KUKA KRL program: MAIN_1.src

&ACCESS RVP
&REL 1
&PARAM TEMPLATE = C:\KRC\Roboter\Template\vorgabe
&PARAM EDITMASK = *
DEF MAIN_1 ( )

; External program calls:
EXT REMOTE_PROG_CALL_171()
EXT PICK_PART_111()
EXT PLACE_PART_112()
EXT EVENT_PROG_START_101()
EXT EVENT_PATH_APPROACH_102()
EXT EVENT_PATH_START_103()
EXT EVENT_PATH_FINISH_105()
EXT EVENT_PATH_RETRACT_106()
EXT EVENT_PROG_FINISH_107()
EXT PROG_1___with_a_very_long_name_and_special_characters()


EXT CLEENING ()
;FOLD INI

;FOLD BASISTECH INI
GLOBAL INTERRUPT DECL 3 WHEN $STOPMESS==TRUE DO IR_STOPM ( )
INTERRUPT ON 3
BAS (#INITMOV,0)
BAS (#VEL_PTP,20)
BAS (#ACC_PTP,20)
;ENDFOLD (BASISTECH INI)

;FOLD SPOTTECH INI
;USERSPOT(#INIT)
;ENDFOLD (SPOTTECH INI)

;FOLD GRIPPERTECH INI
;USER_GRP(0,DUMMY,DUMMY,GDEFAULT)
;ENDFOLD (GRIPPERTECH INI)

;FOLD ARCTECHDIGITAL INI
IF ARC20==TRUE THEN
  A20 (ARC_INI)
  INTERRUPT DECL 6 WHEN $CYCFLAG[3]==FALSE DO A20(TECH_STOP2)
ENDIF
;ENDFOLD (ARCTECHDIGITAL INI)

;FOLD USER INI
;---- Make your modifications here ----

;ENDFOLD (USER INI)

;ENDFOLD (INI)


;FOLD PTP HOME Vel=20 % DEFAULT;%{PE}%R 5.6.13,%MKUKATPBASIS,%CMOVE,%VPTP,%P 1:PTP, 2:HOME, 3:, 5:20, 7:DEFAULT
$BWDSTART=FALSE
PDAT_ACT=PDEFAULT
FDAT_ACT=FHOME
BAS(#PTP_PARAMS,20)
$H_POS=XHOME
PTP XHOME
;ENDFOLD


; Program generated by RoboDK v5.6.9 for RoboDK Industrial on 26/02/2024 09:58:20
; Using nominal kinematics.
;FOLD PTP P1 Vel=100.000 % PDAT1 Tool[1] Base[1];%{PE}%R 5.5.31,%MKUKATPBASIS,%CMOVE,%VPTP,%P 1:PTP, 2:P1, 3:, 5:100.000, 7:PDAT1
$BWDSTART=FALSE
PDAT_ACT=PPDAT1
FDAT_ACT=FP1
BAS(#PTP_PARAMS,100)
PTP XP1 C_PTP
;ENDFOLD

;FOLD PTP P2 Vel=100.000 % PDAT2 Tool[1] Base[1];%{PE}%R 5.5.31,%MKUKATPBASIS,%CMOVE,%VPTP,%P 1:PTP, 2:P2, 3:, 5:100.000, 7:PDAT2
$BWDSTART=FALSE
PDAT_ACT=PPDAT2
FDAT_ACT=FP2
BAS(#PTP_PARAMS,100)
PTP XP2 C_PTP
;ENDFOLD

;FOLD LIN P3 Vel=1.000 m/s CPDAT3 Tool[1] Base[1];%{PE}%R 5.5.0,%MKUKATPA20,%CARC_SWI,%VLIN,%P 1:LIN, 2:P3, 3:, 5:1.000, 7:CPDAT3
$BWDSTART=FALSE
LDAT_ACT=LCPDAT3
FDAT_ACT=FP3
LIN XP3
;ENDFOLD

$OUT[5]=TRUE
$OUT[5]=TRUE
$OUT[5]=0.5
$OUT[5]=true
$ANOUT[5]=TRUE
$ANOUT[5]=TRUE
$ANOUT[5]=0.5
$ANOUT[5]=true
var=val
var=val
WAIT FOR ($IN[5]==TRUE)
WAIT FOR ($IN[5]==TRUE)
WAIT FOR ($IN[5]==0.5)
WAIT FOR ($IN[5]==true)
START_TIMER:
$TIMER_STOP[1]=TRUE
$TIMER_FLAG[1]=FALSE
$TIMER[1]=0.100
$TIMER_STOP[1]=FALSE
WAIT FOR ($IN[5]==TRUE OR $TIMER_FLAG[1])
$TIMER_STOP[1]=TRUE
IF $TIMER_FLAG[1]== TRUE THEN
    HALT ; Timed out!
    GOTO START_TIMER
ENDIF
WAIT FOR (var==val)
START_TIMER:
$TIMER_STOP[1]=TRUE
$TIMER_FLAG[1]=FALSE
$TIMER[1]=0.100
$TIMER_STOP[1]=FALSE
WAIT FOR (var==val OR $TIMER_FLAG[1])
$TIMER_STOP[1]=TRUE
IF $TIMER_FLAG[1]== TRUE THEN
    HALT ; Timed out!
    GOTO START_TIMER
ENDIF
Wait for StrClear($LOOP_MSG[])
$LOOP_CONT = TRUE
$LOOP_MSG[] = "Message"
REMOTE_PROG_CALL_171()
CODE_INSERT_172
; Insert Comment
BASE_DATA[1] = {FRAME: X 719.013,Y -664.003,Z 0.000,A 0.000,B 0.000,C 0.000}
TOOL_DATA[1] = {FRAME: X 129.073,Y 0.000,Z 85.477,A 0.000,B 22.849,C 0.000}
$ACC.ORI1 = 800.00000
$ACC.ORI2 = 800.00000
$VEL.ORI1 = 500.00000
$VEL.ORI2 = 500.00000
$APO.CPTP = 10
$APO.CDIS = 10.000
;FOLD PTP P4 CONT Vel=100.000 % PDAT4 Tool[1] Base[1];%{PE}%R 5.5.31,%MKUKATPBASIS,%CMOVE,%VPTP,%P 1:PTP, 2:P4, 3:C_PTP, 5:100.000, 7:PDAT4
$BWDSTART=FALSE
PDAT_ACT=PPDAT4
FDAT_ACT=FP4
BAS(#PTP_PARAMS,100)
PTP XP4 C_PTP
;ENDFOLD

$ACC.CP = 0.20000
;FOLD LIN P5 Vel=0.100 m/s CPDAT5 Tool[1] Base[1];%{PE}%R 5.5.0,%MKUKATPA20,%CARC_SWI,%VLIN,%P 1:LIN, 2:P5, 3:, 5:0.100, 7:CPDAT5
$BWDSTART=FALSE
LDAT_ACT=LCPDAT5
FDAT_ACT=FP5
LIN XP5
;ENDFOLD

$OUT[5]=TRUE
PICK_PART_111()
$APO.CPTP = 10
$APO.CDIS = 10.000
$ACC.CP = 0.60000
; Linear movement using joint targets is not supported. Change the target type to cartesian or use a joint movement.
;FOLD LIN P6 CONT Vel=0.300 m/s CPDAT6 Tool[1] Base[1];%{PE}%R 5.5.0,%MKUKATPA20,%CARC_SWI,%VLIN,%P 1:LIN, 2:P6, 3:C_DIS, 5:0.300, 7:CPDAT6
$BWDSTART=FALSE
LDAT_ACT=LCPDAT6
FDAT_ACT=FP6
LIN XP6 C_DIS
;ENDFOLD

$ACC.CP = 0.20000
; MoveSearch command not implemented
;FOLD LIN P7 Vel=0.100 m/s CPDAT7 Tool[1] Base[1];%{PE}%R 5.5.0,%MKUKATPA20,%CARC_SWI,%VLIN,%P 1:LIN, 2:P7, 3:, 5:0.100, 7:CPDAT7
$BWDSTART=FALSE
LDAT_ACT=LCPDAT7
FDAT_ACT=FP7
LIN XP7
;ENDFOLD

$OUT[5]=FALSE
PLACE_PART_112()
$APO.CPTP = 10
$APO.CDIS = 10.000
;FOLD LIN P8 CONT Vel=0.100 m/s CPDAT8 Tool[1] Base[1];%{PE}%R 5.5.0,%MKUKATPA20,%CARC_SWI,%VLIN,%P 1:LIN, 2:P8, 3:C_DIS, 5:0.100, 7:CPDAT8
$BWDSTART=FALSE
LDAT_ACT=LCPDAT8
FDAT_ACT=FP8
LIN XP8 C_DIS
;ENDFOLD

BASE_DATA[1] = {FRAME: X 577.670,Y 392.250,Z 0.000,A 38.960,B 0.000,C 0.000}
$APO.CPTP = 25
$APO.CDIS = 25.000
$ACC.ORI1 = 800.00000
$ACC.ORI2 = 800.00000
$VEL.ORI1 = 500.00000
$VEL.ORI2 = 500.00000
$ACC.CP = 0.20000
;FOLD PTP P9 CONT Vel=100.000 % PDAT9 Tool[1] Base[1];%{PE}%R 5.5.31,%MKUKATPBASIS,%CMOVE,%VPTP,%P 1:PTP, 2:P9, 3:C_PTP, 5:100.000, 7:PDAT9
$BWDSTART=FALSE
PDAT_ACT=PPDAT9
FDAT_ACT=FP9
BAS(#PTP_PARAMS,100)
PTP XP9 C_PTP
;ENDFOLD

CIRC {X 430.047,Y 43.774,Z 231.503,A -134.549,B 11.181,C 178.913},{X 109.688,Y -153.222,Z 161.073,A -134.549,B 11.181,C 178.913} C_DIS
; Circular movement using joint targets is not supported. Change the target type to cartesian or use a joint movement.
$ACC.CP = 0.20000
;FOLD LIN P10 Vel=0.100 m/s CPDAT10 Tool[1] Base[1];%{PE}%R 5.5.0,%MKUKATPA20,%CARC_SWI,%VLIN,%P 1:LIN, 2:P10, 3:, 5:0.100, 7:CPDAT10
$BWDSTART=FALSE
LDAT_ACT=LCPDAT10
FDAT_ACT=FP10
LIN XP10
;ENDFOLD

;FOLD PTP P11 Vel=100.000 % PDAT11 Tool[1] Base[1];%{PE}%R 5.5.31,%MKUKATPBASIS,%CMOVE,%VPTP,%P 1:PTP, 2:P11, 3:, 5:100.000, 7:PDAT11
$BWDSTART=FALSE
PDAT_ACT=PPDAT11
FDAT_ACT=FP11
BAS(#PTP_PARAMS,100)
PTP XP11 C_PTP
;ENDFOLD

BASE_DATA[1] = {FRAME: X 0.000,Y 782.714,Z 377.610,A 0.000,B 0.000,C 0.000}
;FOLD PTP P12 Vel=100.000 % PDAT12 Tool[1] Base[1];%{PE}%R 5.5.31,%MKUKATPBASIS,%CMOVE,%VPTP,%P 1:PTP, 2:P12, 3:, 5:100.000, 7:PDAT12
$BWDSTART=FALSE
PDAT_ACT=PPDAT12
FDAT_ACT=FP12
BAS(#PTP_PARAMS,100)
PTP XP12 C_PTP
;ENDFOLD

;FOLD LIN P13 Vel=0.100 m/s CPDAT13 Tool[1] Base[1];%{PE}%R 5.5.0,%MKUKATPA20,%CARC_SWI,%VLIN,%P 1:LIN, 2:P13, 3:, 5:0.100, 7:CPDAT13
$BWDSTART=FALSE
LDAT_ACT=LCPDAT13
FDAT_ACT=FP13
LIN XP13
;ENDFOLD

;FOLD LIN P14 Vel=0.100 m/s CPDAT14 Tool[1] Base[1];%{PE}%R 5.5.0,%MKUKATPA20,%CARC_SWI,%VLIN,%P 1:LIN, 2:P14, 3:, 5:0.100, 7:CPDAT14
$BWDSTART=FALSE
LDAT_ACT=LCPDAT14
FDAT_ACT=FP14
LIN XP14
;ENDFOLD

;FOLD LIN P15 Vel=0.100 m/s CPDAT15 Tool[1] Base[1];%{PE}%R 5.5.0,%MKUKATPA20,%CARC_SWI,%VLIN,%P 1:LIN, 2:P15, 3:, 5:0.100, 7:CPDAT15
$BWDSTART=FALSE
LDAT_ACT=LCPDAT15
FDAT_ACT=FP15
LIN XP15
;ENDFOLD

;FOLD LIN P16 Vel=0.100 m/s CPDAT16 Tool[1] Base[1];%{PE}%R 5.5.0,%MKUKATPA20,%CARC_SWI,%VLIN,%P 1:LIN, 2:P16, 3:, 5:0.100, 7:CPDAT16
$BWDSTART=FALSE
LDAT_ACT=LCPDAT16
FDAT_ACT=FP16
LIN XP16
;ENDFOLD

;FOLD LIN P17 Vel=0.100 m/s CPDAT17 Tool[1] Base[1];%{PE}%R 5.5.0,%MKUKATPA20,%CARC_SWI,%VLIN,%P 1:LIN, 2:P17, 3:, 5:0.100, 7:CPDAT17
$BWDSTART=FALSE
LDAT_ACT=LCPDAT17
FDAT_ACT=FP17
LIN XP17
;ENDFOLD

;FOLD LIN P18 Vel=0.100 m/s CPDAT18 Tool[1] Base[1];%{PE}%R 5.5.0,%MKUKATPA20,%CARC_SWI,%VLIN,%P 1:LIN, 2:P18, 3:, 5:0.100, 7:CPDAT18
$BWDSTART=FALSE
LDAT_ACT=LCPDAT18
FDAT_ACT=FP18
LIN XP18
;ENDFOLD

;FOLD LIN P19 Vel=0.100 m/s CPDAT19 Tool[1] Base[1];%{PE}%R 5.5.0,%MKUKATPA20,%CARC_SWI,%VLIN,%P 1:LIN, 2:P19, 3:, 5:0.100, 7:CPDAT19
$BWDSTART=FALSE
LDAT_ACT=LCPDAT19
FDAT_ACT=FP19
LIN XP19
;ENDFOLD

;FOLD PTP P20 Vel=100.000 % PDAT20 Tool[1] Base[1];%{PE}%R 5.5.31,%MKUKATPBASIS,%CMOVE,%VPTP,%P 1:PTP, 2:P20, 3:, 5:100.000, 7:PDAT20
$BWDSTART=FALSE
PDAT_ACT=PPDAT20
FDAT_ACT=FP20
BAS(#PTP_PARAMS,100)
PTP XP20 C_PTP
;ENDFOLD

EVENT_PROG_START_101()
$APO.CPTP = 1
$APO.CDIS = 1.000
BASE_DATA[1] = {FRAME: X 13.637,Y -840.080,Z 0.000,A -90.000,B 0.000,C 0.000}
; Show Tool 1
;FOLD PTP P21 CONT Vel=100.000 % PDAT21 Tool[1] Base[1];%{PE}%R 5.5.31,%MKUKATPBASIS,%CMOVE,%VPTP,%P 1:PTP, 2:P21, 3:C_PTP, 5:100.000, 7:PDAT21
$BWDSTART=FALSE
PDAT_ACT=PPDAT21
FDAT_ACT=FP21
BAS(#PTP_PARAMS,100)
PTP XP21 C_PTP
;ENDFOLD

EVENT_PATH_APPROACH_102()
;FOLD LIN P22 CONT Vel=1.000 m/s CPDAT22 Tool[1] Base[1];%{PE}%R 5.5.0,%MKUKATPA20,%CARC_SWI,%VLIN,%P 1:LIN, 2:P22, 3:C_DIS, 5:1.000, 7:CPDAT22
$BWDSTART=FALSE
LDAT_ACT=LCPDAT22
FDAT_ACT=FP22
LIN XP22 C_DIS
;ENDFOLD

;FOLD LIN P23 CONT Vel=1.000 m/s CPDAT23 Tool[1] Base[1];%{PE}%R 5.5.0,%MKUKATPA20,%CARC_SWI,%VLIN,%P 1:LIN, 2:P23, 3:C_DIS, 5:1.000, 7:CPDAT23
$BWDSTART=FALSE
LDAT_ACT=LCPDAT23
FDAT_ACT=FP23
LIN XP23 C_DIS
;ENDFOLD

EVENT_PATH_START_103()
;FOLD LIN P24 CONT Vel=0.050 m/s CPDAT24 Tool[1] Base[1];%{PE}%R 5.5.0,%MKUKATPA20,%CARC_SWI,%VLIN,%P 1:LIN, 2:P24, 3:C_DIS, 5:0.050, 7:CPDAT24
$BWDSTART=FALSE
LDAT_ACT=LCPDAT24
FDAT_ACT=FP24
LIN XP24 C_DIS
;ENDFOLD

;FOLD LIN P25 CONT Vel=0.050 m/s CPDAT25 Tool[1] Base[1];%{PE}%R 5.5.0,%MKUKATPA20,%CARC_SWI,%VLIN,%P 1:LIN, 2:P25, 3:C_DIS, 5:0.050, 7:CPDAT25
$BWDSTART=FALSE
LDAT_ACT=LCPDAT25
FDAT_ACT=FP25
LIN XP25 C_DIS
;ENDFOLD

;FOLD LIN P26 CONT Vel=0.050 m/s CPDAT26 Tool[1] Base[1];%{PE}%R 5.5.0,%MKUKATPA20,%CARC_SWI,%VLIN,%P 1:LIN, 2:P26, 3:C_DIS, 5:0.050, 7:CPDAT26
$BWDSTART=FALSE
LDAT_ACT=LCPDAT26
FDAT_ACT=FP26
LIN XP26 C_DIS
;ENDFOLD

;FOLD LIN P27 CONT Vel=0.050 m/s CPDAT27 Tool[1] Base[1];%{PE}%R 5.5.0,%MKUKATPA20,%CARC_SWI,%VLIN,%P 1:LIN, 2:P27, 3:C_DIS, 5:0.050, 7:CPDAT27
$BWDSTART=FALSE
LDAT_ACT=LCPDAT27
FDAT_ACT=FP27
LIN XP27 C_DIS
;ENDFOLD

;FOLD LIN P28 CONT Vel=0.050 m/s CPDAT28 Tool[1] Base[1];%{PE}%R 5.5.0,%MKUKATPA20,%CARC_SWI,%VLIN,%P 1:LIN, 2:P28, 3:C_DIS, 5:0.050, 7:CPDAT28
$BWDSTART=FALSE
LDAT_ACT=LCPDAT28
FDAT_ACT=FP28
LIN XP28 C_DIS
;ENDFOLD

;FOLD LIN P29 CONT Vel=0.050 m/s CPDAT29 Tool[1] Base[1];%{PE}%R 5.5.0,%MKUKATPA20,%CARC_SWI,%VLIN,%P 1:LIN, 2:P29, 3:C_DIS, 5:0.050, 7:CPDAT29
$BWDSTART=FALSE
LDAT_ACT=LCPDAT29
FDAT_ACT=FP29
LIN XP29 C_DIS
;ENDFOLD

;FOLD LIN P30 CONT Vel=0.050 m/s CPDAT30 Tool[1] Base[1];%{PE}%R 5.5.0,%MKUKATPA20,%CARC_SWI,%VLIN,%P 1:LIN, 2:P30, 3:C_DIS, 5:0.050, 7:CPDAT30
$BWDSTART=FALSE
LDAT_ACT=LCPDAT30
FDAT_ACT=FP30
LIN XP30 C_DIS
;ENDFOLD

;FOLD LIN P31 CONT Vel=0.050 m/s CPDAT31 Tool[1] Base[1];%{PE}%R 5.5.0,%MKUKATPA20,%CARC_SWI,%VLIN,%P 1:LIN, 2:P31, 3:C_DIS, 5:0.050, 7:CPDAT31
$BWDSTART=FALSE
LDAT_ACT=LCPDAT31
FDAT_ACT=FP31
LIN XP31 C_DIS
;ENDFOLD

;FOLD LIN P32 CONT Vel=0.050 m/s CPDAT32 Tool[1] Base[1];%{PE}%R 5.5.0,%MKUKATPA20,%CARC_SWI,%VLIN,%P 1:LIN, 2:P32, 3:C_DIS, 5:0.050, 7:CPDAT32
$BWDSTART=FALSE
LDAT_ACT=LCPDAT32
FDAT_ACT=FP32
LIN XP32 C_DIS
;ENDFOLD

;FOLD LIN P33 CONT Vel=0.050 m/s CPDAT33 Tool[1] Base[1];%{PE}%R 5.5.0,%MKUKATPA20,%CARC_SWI,%VLIN,%P 1:LIN, 2:P33, 3:C_DIS, 5:0.050, 7:CPDAT33
$BWDSTART=FALSE
LDAT_ACT=LCPDAT33
FDAT_ACT=FP33
LIN XP33 C_DIS
;ENDFOLD

;FOLD LIN P34 CONT Vel=0.050 m/s CPDAT34 Tool[1] Base[1];%{PE}%R 5.5.0,%MKUKATPA20,%CARC_SWI,%VLIN,%P 1:LIN, 2:P34, 3:C_DIS, 5:0.050, 7:CPDAT34
$BWDSTART=FALSE
LDAT_ACT=LCPDAT34
FDAT_ACT=FP34
LIN XP34 C_DIS
;ENDFOLD

;FOLD LIN P35 CONT Vel=0.050 m/s CPDAT35 Tool[1] Base[1];%{PE}%R 5.5.0,%MKUKATPA20,%CARC_SWI,%VLIN,%P 1:LIN, 2:P35, 3:C_DIS, 5:0.050, 7:CPDAT35
$BWDSTART=FALSE
LDAT_ACT=LCPDAT35
FDAT_ACT=FP35
LIN XP35 C_DIS
;ENDFOLD

;FOLD LIN P36 CONT Vel=0.050 m/s CPDAT36 Tool[1] Base[1];%{PE}%R 5.5.0,%MKUKATPA20,%CARC_SWI,%VLIN,%P 1:LIN, 2:P36, 3:C_DIS, 5:0.050, 7:CPDAT36
$BWDSTART=FALSE
LDAT_ACT=LCPDAT36
FDAT_ACT=FP36
LIN XP36 C_DIS
;ENDFOLD

;FOLD LIN P37 CONT Vel=0.050 m/s CPDAT37 Tool[1] Base[1];%{PE}%R 5.5.0,%MKUKATPA20,%CARC_SWI,%VLIN,%P 1:LIN, 2:P37, 3:C_DIS, 5:0.050, 7:CPDAT37
$BWDSTART=FALSE
LDAT_ACT=LCPDAT37
FDAT_ACT=FP37
LIN XP37 C_DIS
;ENDFOLD

;FOLD LIN P38 CONT Vel=0.050 m/s CPDAT38 Tool[1] Base[1];%{PE}%R 5.5.0,%MKUKATPA20,%CARC_SWI,%VLIN,%P 1:LIN, 2:P38, 3:C_DIS, 5:0.050, 7:CPDAT38
$BWDSTART=FALSE
LDAT_ACT=LCPDAT38
FDAT_ACT=FP38
LIN XP38 C_DIS
;ENDFOLD

;FOLD LIN P39 CONT Vel=0.050 m/s CPDAT39 Tool[1] Base[1];%{PE}%R 5.5.0,%MKUKATPA20,%CARC_SWI,%VLIN,%P 1:LIN, 2:P39, 3:C_DIS, 5:0.050, 7:CPDAT39
$BWDSTART=FALSE
LDAT_ACT=LCPDAT39
FDAT_ACT=FP39
LIN XP39 C_DIS
;ENDFOLD

;FOLD LIN P40 CONT Vel=0.050 m/s CPDAT40 Tool[1] Base[1];%{PE}%R 5.5.0,%MKUKATPA20,%CARC_SWI,%VLIN,%P 1:LIN, 2:P40, 3:C_DIS, 5:0.050, 7:CPDAT40
$BWDSTART=FALSE
LDAT_ACT=LCPDAT40
FDAT_ACT=FP40
LIN XP40 C_DIS
;ENDFOLD

;FOLD LIN P41 CONT Vel=0.050 m/s CPDAT41 Tool[1] Base[1];%{PE}%R 5.5.0,%MKUKATPA20,%CARC_SWI,%VLIN,%P 1:LIN, 2:P41, 3:C_DIS, 5:0.050, 7:CPDAT41
$BWDSTART=FALSE
LDAT_ACT=LCPDAT41
FDAT_ACT=FP41
LIN XP41 C_DIS
;ENDFOLD

;FOLD LIN P42 CONT Vel=0.050 m/s CPDAT42 Tool[1] Base[1];%{PE}%R 5.5.0,%MKUKATPA20,%CARC_SWI,%VLIN,%P 1:LIN, 2:P42, 3:C_DIS, 5:0.050, 7:CPDAT42
$BWDSTART=FALSE
LDAT_ACT=LCPDAT42
FDAT_ACT=FP42
LIN XP42 C_DIS
;ENDFOLD

;FOLD LIN P43 CONT Vel=0.050 m/s CPDAT43 Tool[1] Base[1];%{PE}%R 5.5.0,%MKUKATPA20,%CARC_SWI,%VLIN,%P 1:LIN, 2:P43, 3:C_DIS, 5:0.050, 7:CPDAT43
$BWDSTART=FALSE
LDAT_ACT=LCPDAT43
FDAT_ACT=FP43
LIN XP43 C_DIS
;ENDFOLD

;FOLD LIN P44 CONT Vel=0.050 m/s CPDAT44 Tool[1] Base[1];%{PE}%R 5.5.0,%MKUKATPA20,%CARC_SWI,%VLIN,%P 1:LIN, 2:P44, 3:C_DIS, 5:0.050, 7:CPDAT44
$BWDSTART=FALSE
LDAT_ACT=LCPDAT44
FDAT_ACT=FP44
LIN XP44 C_DIS
;ENDFOLD

;FOLD LIN P45 CONT Vel=0.050 m/s CPDAT45 Tool[1] Base[1];%{PE}%R 5.5.0,%MKUKATPA20,%CARC_SWI,%VLIN,%P 1:LIN, 2:P45, 3:C_DIS, 5:0.050, 7:CPDAT45
$BWDSTART=FALSE
LDAT_ACT=LCPDAT45
FDAT_ACT=FP45
LIN XP45 C_DIS
;ENDFOLD

;FOLD LIN P46 CONT Vel=0.050 m/s CPDAT46 Tool[1] Base[1];%{PE}%R 5.5.0,%MKUKATPA20,%CARC_SWI,%VLIN,%P 1:LIN, 2:P46, 3:C_DIS, 5:0.050, 7:CPDAT46
$BWDSTART=FALSE
LDAT_ACT=LCPDAT46
FDAT_ACT=FP46
LIN XP46 C_DIS
;ENDFOLD

;FOLD LIN P47 CONT Vel=0.050 m/s CPDAT47 Tool[1] Base[1];%{PE}%R 5.5.0,%MKUKATPA20,%CARC_SWI,%VLIN,%P 1:LIN, 2:P47, 3:C_DIS, 5:0.050, 7:CPDAT47
$BWDSTART=FALSE
LDAT_ACT=LCPDAT47
FDAT_ACT=FP47
LIN XP47 C_DIS
;ENDFOLD

;FOLD LIN P48 CONT Vel=0.050 m/s CPDAT48 Tool[1] Base[1];%{PE}%R 5.5.0,%MKUKATPA20,%CARC_SWI,%VLIN,%P 1:LIN, 2:P48, 3:C_DIS, 5:0.050, 7:CPDAT48
$BWDSTART=FALSE
LDAT_ACT=LCPDAT48
FDAT_ACT=FP48
LIN XP48 C_DIS
;ENDFOLD

;FOLD LIN P49 CONT Vel=0.050 m/s CPDAT49 Tool[1] Base[1];%{PE}%R 5.5.0,%MKUKATPA20,%CARC_SWI,%VLIN,%P 1:LIN, 2:P49, 3:C_DIS, 5:0.050, 7:CPDAT49
$BWDSTART=FALSE
LDAT_ACT=LCPDAT49
FDAT_ACT=FP49
LIN XP49 C_DIS
;ENDFOLD

;FOLD LIN P50 CONT Vel=0.050 m/s CPDAT50 Tool[1] Base[1];%{PE}%R 5.5.0,%MKUKATPA20,%CARC_SWI,%VLIN,%P 1:LIN, 2:P50, 3:C_DIS, 5:0.050, 7:CPDAT50
$BWDSTART=FALSE
LDAT_ACT=LCPDAT50
FDAT_ACT=FP50
LIN XP50 C_DIS
;ENDFOLD

;FOLD LIN P51 CONT Vel=0.050 m/s CPDAT51 Tool[1] Base[1];%{PE}%R 5.5.0,%MKUKATPA20,%CARC_SWI,%VLIN,%P 1:LIN, 2:P51, 3:C_DIS, 5:0.050, 7:CPDAT51
$BWDSTART=FALSE
LDAT_ACT=LCPDAT51
FDAT_ACT=FP51
LIN XP51 C_DIS
;ENDFOLD

;FOLD LIN P52 CONT Vel=0.050 m/s CPDAT52 Tool[1] Base[1];%{PE}%R 5.5.0,%MKUKATPA20,%CARC_SWI,%VLIN,%P 1:LIN, 2:P52, 3:C_DIS, 5:0.050, 7:CPDAT52
$BWDSTART=FALSE
LDAT_ACT=LCPDAT52
FDAT_ACT=FP52
LIN XP52 C_DIS
;ENDFOLD

;FOLD LIN P53 CONT Vel=0.050 m/s CPDAT53 Tool[1] Base[1];%{PE}%R 5.5.0,%MKUKATPA20,%CARC_SWI,%VLIN,%P 1:LIN, 2:P53, 3:C_DIS, 5:0.050, 7:CPDAT53
$BWDSTART=FALSE
LDAT_ACT=LCPDAT53
FDAT_ACT=FP53
LIN XP53 C_DIS
;ENDFOLD

;FOLD LIN P54 CONT Vel=0.050 m/s CPDAT54 Tool[1] Base[1];%{PE}%R 5.5.0,%MKUKATPA20,%CARC_SWI,%VLIN,%P 1:LIN, 2:P54, 3:C_DIS, 5:0.050, 7:CPDAT54
$BWDSTART=FALSE
LDAT_ACT=LCPDAT54
FDAT_ACT=FP54
LIN XP54 C_DIS
;ENDFOLD

;FOLD LIN P55 CONT Vel=0.050 m/s CPDAT55 Tool[1] Base[1];%{PE}%R 5.5.0,%MKUKATPA20,%CARC_SWI,%VLIN,%P 1:LIN, 2:P55, 3:C_DIS, 5:0.050, 7:CPDAT55
$BWDSTART=FALSE
LDAT_ACT=LCPDAT55
FDAT_ACT=FP55
LIN XP55 C_DIS
;ENDFOLD

;FOLD LIN P56 CONT Vel=0.050 m/s CPDAT56 Tool[1] Base[1];%{PE}%R 5.5.0,%MKUKATPA20,%CARC_SWI,%VLIN,%P 1:LIN, 2:P56, 3:C_DIS, 5:0.050, 7:CPDAT56
$BWDSTART=FALSE
LDAT_ACT=LCPDAT56
FDAT_ACT=FP56
LIN XP56 C_DIS
;ENDFOLD

;FOLD LIN P57 CONT Vel=0.050 m/s CPDAT57 Tool[1] Base[1];%{PE}%R 5.5.0,%MKUKATPA20,%CARC_SWI,%VLIN,%P 1:LIN, 2:P57, 3:C_DIS, 5:0.050, 7:CPDAT57
$BWDSTART=FALSE
LDAT_ACT=LCPDAT57
FDAT_ACT=FP57
LIN XP57 C_DIS
;ENDFOLD

;FOLD LIN P58 CONT Vel=0.050 m/s CPDAT58 Tool[1] Base[1];%{PE}%R 5.5.0,%MKUKATPA20,%CARC_SWI,%VLIN,%P 1:LIN, 2:P58, 3:C_DIS, 5:0.050, 7:CPDAT58
$BWDSTART=FALSE
LDAT_ACT=LCPDAT58
FDAT_ACT=FP58
LIN XP58 C_DIS
;ENDFOLD

;FOLD LIN P59 CONT Vel=0.050 m/s CPDAT59 Tool[1] Base[1];%{PE}%R 5.5.0,%MKUKATPA20,%CARC_SWI,%VLIN,%P 1:LIN, 2:P59, 3:C_DIS, 5:0.050, 7:CPDAT59
$BWDSTART=FALSE
LDAT_ACT=LCPDAT59
FDAT_ACT=FP59
LIN XP59 C_DIS
;ENDFOLD

;FOLD LIN P60 CONT Vel=0.050 m/s CPDAT60 Tool[1] Base[1];%{PE}%R 5.5.0,%MKUKATPA20,%CARC_SWI,%VLIN,%P 1:LIN, 2:P60, 3:C_DIS, 5:0.050, 7:CPDAT60
$BWDSTART=FALSE
LDAT_ACT=LCPDAT60
FDAT_ACT=FP60
LIN XP60 C_DIS
;ENDFOLD

;FOLD LIN P61 CONT Vel=0.050 m/s CPDAT61 Tool[1] Base[1];%{PE}%R 5.5.0,%MKUKATPA20,%CARC_SWI,%VLIN,%P 1:LIN, 2:P61, 3:C_DIS, 5:0.050, 7:CPDAT61
$BWDSTART=FALSE
LDAT_ACT=LCPDAT61
FDAT_ACT=FP61
LIN XP61 C_DIS
;ENDFOLD

;FOLD LIN P62 CONT Vel=0.050 m/s CPDAT62 Tool[1] Base[1];%{PE}%R 5.5.0,%MKUKATPA20,%CARC_SWI,%VLIN,%P 1:LIN, 2:P62, 3:C_DIS, 5:0.050, 7:CPDAT62
$BWDSTART=FALSE
LDAT_ACT=LCPDAT62
FDAT_ACT=FP62
LIN XP62 C_DIS
;ENDFOLD

;FOLD LIN P63 CONT Vel=0.050 m/s CPDAT63 Tool[1] Base[1];%{PE}%R 5.5.0,%MKUKATPA20,%CARC_SWI,%VLIN,%P 1:LIN, 2:P63, 3:C_DIS, 5:0.050, 7:CPDAT63
$BWDSTART=FALSE
LDAT_ACT=LCPDAT63
FDAT_ACT=FP63
LIN XP63 C_DIS
;ENDFOLD

;FOLD LIN P64 CONT Vel=0.050 m/s CPDAT64 Tool[1] Base[1];%{PE}%R 5.5.0,%MKUKATPA20,%CARC_SWI,%VLIN,%P 1:LIN, 2:P64, 3:C_DIS, 5:0.050, 7:CPDAT64
$BWDSTART=FALSE
LDAT_ACT=LCPDAT64
FDAT_ACT=FP64
LIN XP64 C_DIS
;ENDFOLD

;FOLD LIN P65 CONT Vel=0.050 m/s CPDAT65 Tool[1] Base[1];%{PE}%R 5.5.0,%MKUKATPA20,%CARC_SWI,%VLIN,%P 1:LIN, 2:P65, 3:C_DIS, 5:0.050, 7:CPDAT65
$BWDSTART=FALSE
LDAT_ACT=LCPDAT65
FDAT_ACT=FP65
LIN XP65 C_DIS
;ENDFOLD

;FOLD LIN P66 CONT Vel=0.050 m/s CPDAT66 Tool[1] Base[1];%{PE}%R 5.5.0,%MKUKATPA20,%CARC_SWI,%VLIN,%P 1:LIN, 2:P66, 3:C_DIS, 5:0.050, 7:CPDAT66
$BWDSTART=FALSE
LDAT_ACT=LCPDAT66
FDAT_ACT=FP66
LIN XP66 C_DIS
;ENDFOLD

;FOLD LIN P67 CONT Vel=0.050 m/s CPDAT67 Tool[1] Base[1];%{PE}%R 5.5.0,%MKUKATPA20,%CARC_SWI,%VLIN,%P 1:LIN, 2:P67, 3:C_DIS, 5:0.050, 7:CPDAT67
$BWDSTART=FALSE
LDAT_ACT=LCPDAT67
FDAT_ACT=FP67
LIN XP67 C_DIS
;ENDFOLD

;FOLD LIN P68 CONT Vel=0.050 m/s CPDAT68 Tool[1] Base[1];%{PE}%R 5.5.0,%MKUKATPA20,%CARC_SWI,%VLIN,%P 1:LIN, 2:P68, 3:C_DIS, 5:0.050, 7:CPDAT68
$BWDSTART=FALSE
LDAT_ACT=LCPDAT68
FDAT_ACT=FP68
LIN XP68 C_DIS
;ENDFOLD

EVENT_PATH_FINISH_105()
;FOLD LIN P69 CONT Vel=1.000 m/s CPDAT69 Tool[1] Base[1];%{PE}%R 5.5.0,%MKUKATPA20,%CARC_SWI,%VLIN,%P 1:LIN, 2:P69, 3:C_DIS, 5:1.000, 7:CPDAT69
$BWDSTART=FALSE
LDAT_ACT=LCPDAT69
FDAT_ACT=FP69
LIN XP69 C_DIS
;ENDFOLD

;FOLD LIN P70 CONT Vel=1.000 m/s CPDAT70 Tool[1] Base[1];%{PE}%R 5.5.0,%MKUKATPA20,%CARC_SWI,%VLIN,%P 1:LIN, 2:P70, 3:C_DIS, 5:1.000, 7:CPDAT70
$BWDSTART=FALSE
LDAT_ACT=LCPDAT70
FDAT_ACT=FP70
LIN XP70 C_DIS
;ENDFOLD

EVENT_PATH_RETRACT_106()
EVENT_PROG_FINISH_107()
BASE_DATA[1] = {FRAME: X 719.013,Y -664.003,Z 0.000,A 0.000,B 0.000,C 0.000}
;FOLD PTP P71 CONT Vel=100.000 % PDAT71 Tool[1] Base[1];%{PE}%R 5.5.31,%MKUKATPBASIS,%CMOVE,%VPTP,%P 1:PTP, 2:P71, 3:C_PTP, 5:100.000, 7:PDAT71
$BWDSTART=FALSE
PDAT_ACT=PPDAT71
FDAT_ACT=FP71
BAS(#PTP_PARAMS,100)
PTP XP71 C_PTP
;ENDFOLD

WAIT SEC 1.250
;FOLD LIN P72 CONT Vel=1.000 m/s CPDAT72 Tool[1] Base[1];%{PE}%R 5.5.0,%MKUKATPA20,%CARC_SWI,%VLIN,%P 1:LIN, 2:P72, 3:C_DIS, 5:1.000, 7:CPDAT72
$BWDSTART=FALSE
LDAT_ACT=LCPDAT72
FDAT_ACT=FP72
LIN XP72 C_DIS
;ENDFOLD

WAIT FOR ($IN[1]==TRUE)
;FOLD LIN P73 CONT Vel=1.000 m/s CPDAT73 Tool[1] Base[1];%{PE}%R 5.5.0,%MKUKATPA20,%CARC_SWI,%VLIN,%P 1:LIN, 2:P73, 3:C_DIS, 5:1.000, 7:CPDAT73
$BWDSTART=FALSE
LDAT_ACT=LCPDAT73
FDAT_ACT=FP73
LIN XP73 C_DIS
;ENDFOLD

PROG_1___with_a_very_long_name_and_special_characters()
END
